Staubli VAL3: settoolmode.pgx

public program settoolmode()
  local num l_i
begin
  $jogMode(3)
   for l_i = 0 to size(sShowType)-1
    sShowType[l_i]=sCartisiam[l_i]
  endFor
end
